// TIA Portal V20 export
// export: Created 2026-10-19T18:06:05.7697074Z, ExportSetting WithDefaults, DisplayName Totally Integrated Automation Portal, DisplayVersion V20 Update 6, DisplayName TIA Portal Openness, DisplayVersion V20 Update 6, DisplayName TIA Portal Version Control Interface, DisplayVersion V20 Update 6, DisplayName SINAMICS Startdrive Advanced, DisplayVersion V20 SP1, DisplayName SINAMICS Startdrive G130, G150, S120, S150, SINAMICS MV, G220, S200, S210, DisplayVersion V20 SP1, DisplayName SINAMICS Startdrive G110M, G120, G120C, G120D, G120P, G115D, DisplayVersion V20 SP1, DisplayName STEP 7 Professional, DisplayVersion V20 Update 6, DisplayName STEP 7 Safety, DisplayVersion V20 Update 2, DisplayName WinCC Basic/Comfort/Advanced, DisplayVersion V20 Update 6, DisplayName WinCC Unified, DisplayVersion V20 Update 6
FUNCTION "Weighing Station FC" : Void   // FC31, SCL
{ S7_Optimized_Access := 'TRUE' }
VERSION : 0.1
// stored: AutoNumber true, IsIECCheckEnabled false, SetENOAutomatically false, UDAEnableTagReadback false
   VAR_INPUT
      Start : Bool;
      MinWeight : Real;
      MaxWeight : Real;
   END_VAR
BEGIN
   "R_TRIG_DB_25"(CLK:=#Start, Q=> "R_Start_WS");

   CASE "State_WS" OF
       0: // IDLE / READY
           "Control_DB"."Weighing Station".Ready := TRUE;
           "Control_DB"."Weighing Station".Running := FALSE;
           IF "R_Start_WS" THEN
               "Control_DB"."Weighing Station".Done := FALSE;
               "Control_DB"."Weighing Station".Valid := FALSE;
               "Control_DB"."Weighing Station".Ready := FALSE;
               "Control_DB"."Weighing Station".Error_ID := 0;
               "State_WS" := 10;
           END_IF;

       10:
           "Control_DB"."Weighing Station".Start := FALSE;
           "Control_DB"."Weighing Station".Running := TRUE;
           IF "Control_DB".PopUp_Cnv[1].Inputs."Lift Up" THEN

               IF NOT "SAI_Cyclic_WeightProc_DB".DataOK THEN
                   "Control_DB"."Weighing Station".Error_ID.%X0 := TRUE;
                   "Control_DB"."Weighing Station".Done := TRUE;
                   "State_WS" := 100;
               ELSE
                   "Control_DB"."Weighing Station".Weight := "SAI_Cyclic_WeightProc_DB".RealTimeWeight;
                   "State_WS" := 20;
               END_IF;
           END_IF;
           "IEC_Timer_0_DB_17".TON(IN:=TRUE,
                                   PT:=t#10S);
           IF "IEC_Timer_0_DB_17".Q THEN
               "IEC_Timer_0_DB_17".TON(IN := FALSE,
                                       PT := t#0S);
               // "Control_DB"."Weighing Station".Done := TRUE;
               "State_WS" := 20;
           END_IF;

       20:
           IF "Control_DB"."Weighing Station".Weight < #MinWeight THEN
               "Control_DB"."Weighing Station".Valid := FALSE;
               // "Control_DB"."Weighing Station".Error_ID.%X1 := TRUE;
           ELSIF "Control_DB"."Weighing Station".Weight > #MaxWeight THEN
               "Control_DB"."Weighing Station".Valid := FALSE;
               // "Control_DB"."Weighing Station".Error_ID.%X2 := TRUE;
           ELSE
               "Control_DB"."Weighing Station".Valid := TRUE;
               "Control_DB"."Weighing Station".Error_ID := 0;
           END_IF;
           "State_WS" := 100;

       100:
           "Control_DB"."Weighing Station".Running := FALSE;
           "Control_DB"."Weighing Station".Done := TRUE;
           "State_WS" := 0;

   END_CASE;

   IF "Reset_All" THEN
       "Control_DB"."Weighing Station".Error_ID := 0;
   END_IF;
END_FUNCTION
